Omron CX-Programmer project NewProject (CX-Programmer 9.50)

# PLC freezer_iiot: CP1L M

## Global symbols (name address type ; comment)
100 CHANNEL  ; 10sec
100.00 BOOL  ; Out1
1800 CHANNEL  ; 3_min
D0 CHANNEL  ; T * 10
D10 CHANNEL  ; Band/2
D11 CHANNEL  ; SP + Band/2
D12 CHANNEL  ; SP - Band/2
D2 CHANNEL  ; SP
D20 CHANNEL  ; presim_HB
D3 CHANNEL  ; Band
D4 CHANNEL  ; Comp_status
D5 CHANNEL  ; PLC heartbeat
D6 CHANNEL  ; sim heartbeat
D7 CHANNEL  ; COM_Fault
T0000 BOOL  ; 3_min
T0001 BOOL  ; 10sec
T0002 BOOL  ; 12min
T0003 BOOL  ; 8min
W0.00 BOOL  ; Compressor
W0.01 BOOL  ; Closed Compressor
W0.02 BOOL  ; comfault
W0.03 BOOL  ; fallback
W0.04 BOOL  ; strat_Timer8Min

## Program NewProgram1 (cyclic task 0)

### Section Section1

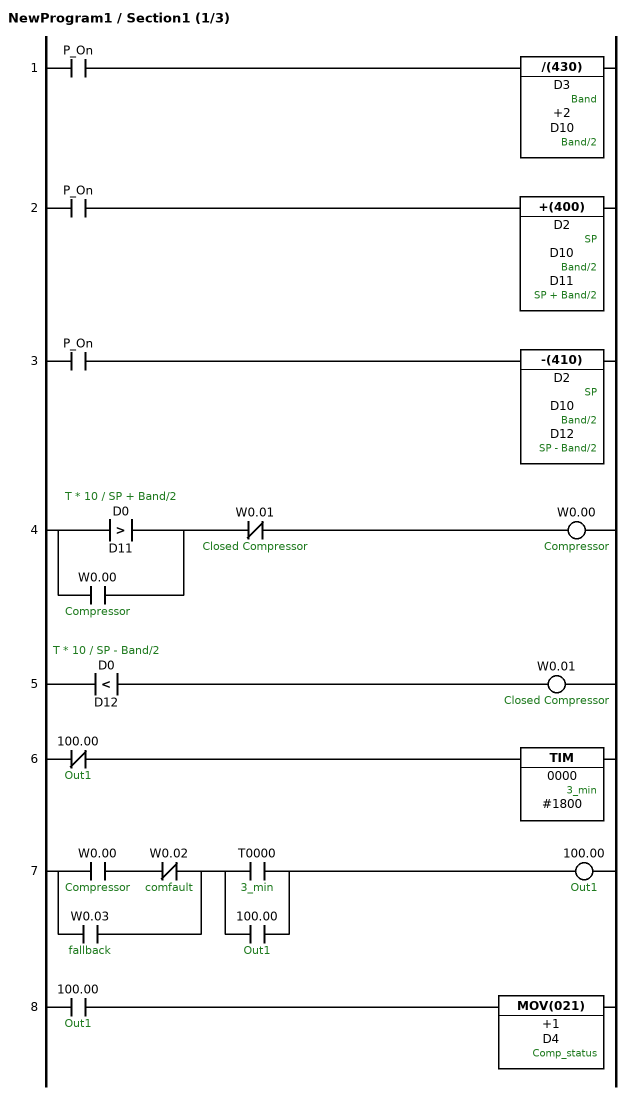
; rung 1
LD P_On
/(430) D3 +2 D10  ; Band, Band/2
; rung 2
LD P_On
+(400) D2 D10 D11  ; SP, Band/2, SP + Band/2
; rung 3
LD P_On
-(410) D2 D10 D12  ; SP, Band/2, SP - Band/2
; rung 4
LD>S(322) D0 D11  ; T * 10, SP + Band/2
OR W0.00  ; Compressor
ANDNOT W0.01  ; Closed Compressor
OUT W0.00  ; Compressor
; rung 5
LD<S(312) D0 D12  ; T * 10, SP - Band/2
OUT W0.01  ; Closed Compressor
; rung 6
LDNOT 100.00  ; Out1
TIM 0000 #1800  ; 3_min
; rung 7
LD W0.00  ; Compressor
ANDNOT W0.02  ; comfault
OR W0.03  ; fallback
LD T0000  ; 3_min
OR 100.00  ; Out1
ANDLD
OUT 100.00  ; Out1
; rung 8
LD 100.00  ; Out1
MOV(021) +1 D4  ; Comp_status

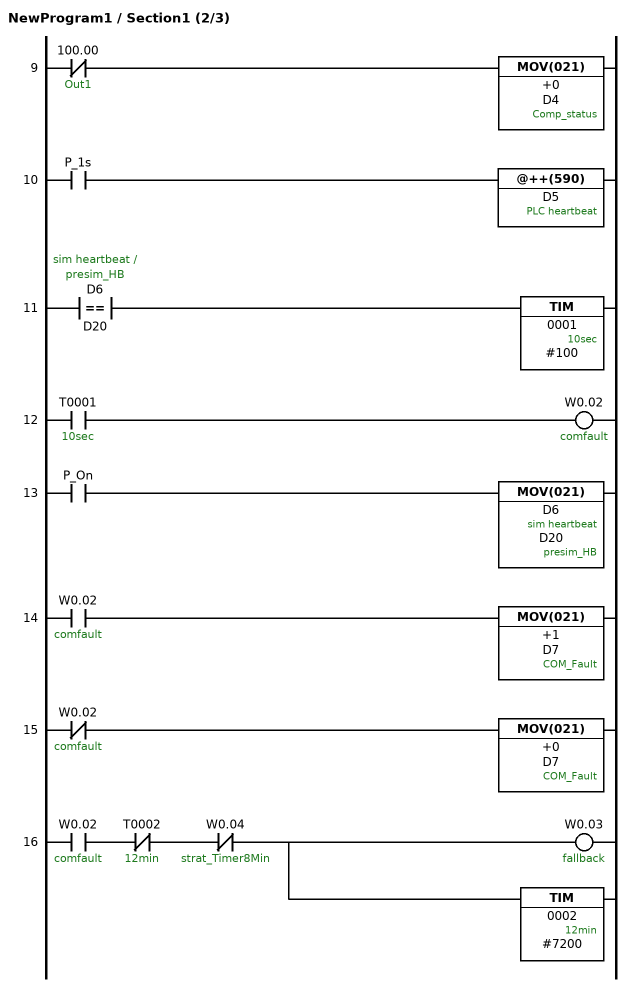
; rung 9
LDNOT 100.00  ; Out1
MOV(021) +0 D4  ; Comp_status
; rung 10
LD P_1s
@++(590) D5  ; PLC heartbeat
; rung 11
LD=(300) D6 D20  ; sim heartbeat, presim_HB
TIM 0001 #100  ; 10sec
; rung 12
LD T0001  ; 10sec
OUT W0.02  ; comfault
; rung 13
LD P_On
MOV(021) D6 D20  ; sim heartbeat, presim_HB
; rung 14
LD W0.02  ; comfault
MOV(021) +1 D7  ; COM_Fault
; rung 15
LDNOT W0.02  ; comfault
MOV(021) +0 D7  ; COM_Fault
; rung 16
LD W0.02  ; comfault
ANDNOT T0002  ; 12min
ANDNOT W0.04  ; strat_Timer8Min
OUT W0.03  ; fallback
TIM 0002 #7200  ; 12min

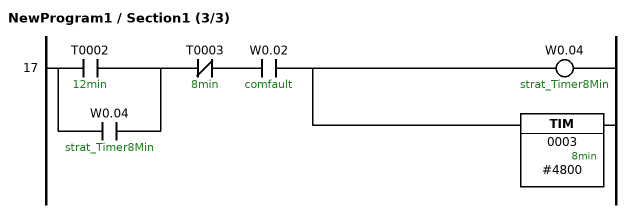
; rung 17
LD T0002  ; 12min
OR W0.04  ; strat_Timer8Min
ANDNOT T0003  ; 8min
AND W0.02  ; comfault
OUT W0.04  ; strat_Timer8Min
TIM 0003 #4800  ; 8min

### Section END
; rung 0
END(001)